// TIA Portal V20 export
Screen "RobotService_Zone05"  1276x673
  ScreenItem "Line_Header_X0_Y64" at 0,64 size 1280x0  Type=HmiLine
  ScreenItem "permanentareaborderrectangle" at 0,0 size 0x0  Type=HmiRectangle
  ScreenItem "Title_ScreenOverview_X390_Y2_3" at 375,5 size 510x57  Type=HmiTextBox
  ScreenItem "190RB04" at 467,72 size 193x297  Type=HmiFaceplateContainer
  ScreenItem "190RB03" at 247,72 size 193x297  Type=HmiFaceplateContainer
  ScreenItem "190" at 27,72 size 189x297  Type=HmiFaceplateContainer
  ScreenItem "Faceplate container_1" at 1127,70 size 127x580  Type=HmiFaceplateContainer
  ScreenItem "Button_Back_1" at 1164,0 size 90x60  Type=HmiButton
  ScreenItem "Button_Back_2" at 8,2 size 90x60  Type=HmiButton
